Fanuc KAREL source: kf00081.KL

-- PROVISIONAL review KL for V1013-1; original PC SHA256 9ff8b2a0835719f867cf2430197b2e038d988fe0204db05fc21fc1ea3921ced4
-- Incomplete behavior may be omitted. Consult companion uncertainty JSON. Do not deploy.
PROGRAM KF00081
%NOLOCKGROUP
BEGIN
  -- UNRESOLVED_PC offsets 5-15; opcodes 27,22,31
  -- UNRESOLVED_PC offsets 20-54; opcodes 27,27,2E,22,22,22,22,31
  -- UNRESOLVED_PC offsets 59-63; opcodes 7F
END KF00081
